Staubli VAL3: ouvrirPince.pgx

program ouvrirPince()
begin
  close(tPince)
end
